Fanuc KAREL source: kx00010.KL

-- PROVISIONAL review KL for V940-1; original PC SHA256 10e6664344693af683a6fdf33c1094fee0b017de838aadd2ae81c3276f144b0f
-- Incomplete behavior may be omitted. Consult companion uncertainty JSON. Do not deploy.
PROGRAM KX00010
%NOLOCKGROUP
VAR
  I : INTEGER
  J : INTEGER
  B : BOOLEAN
  F : FILE
  S : STRING[80]
-- UNRESOLVED_DECL P type=000102
BEGIN
  -- V9_ZERO_TABLE_METADATA_HINT layout=0001; no indexed target words; source/name/runtime held
  -- UNRESOLVED_PC offsets 5-7; opcodes 9C,10
  -- UNRESOLVED_PC offsets 12-16; opcodes 7F
END KX00010
